(*
SPDX-License-Identifier: MIT
License: https://opensource.org/license/mit
*)

(*!
<summary>Owns two ordered single-cycle tests for topology regressions.</summary>
<description>
Owns persistent child storage and fixed parent associations. Use in one task without reentry.
Children is borrowed and must not be modified by application code. Constructor callbacks are not used.
Regression tests may deliberately corrupt the exposed array between failed operations to inject topology faults.
</description>
*)

{attribute 'no_assign'}
{attribute 'no_explicit_call' := 'do not call this function block directly'}
FUNCTION_BLOCK PairTestGroup EXTENDS TOF_Testing.TestGroup<2>
VAR_STAT
	//! <summary>Class name shared by all instances of this function block.</summary>
	{attribute 'hide'}
	_ClassName : STRING := __POUNAME();
END_VAR
VAR
	{attribute 'hide'}
	{attribute 'init_namespace'}
	_NamespaceName : STRING;
END_VAR
VAR_OUTPUT
	//! <summary>First owned regression leaf.</summary>
	First : TestingProbe(name := "First", parent := THIS^);
	//! <summary>Second owned regression leaf.</summary>
	Second : TestingProbe(name := "Second", parent := THIS^);
END_VAR
VAR
	_Children : ARRAY [0.._ChildCount - 1] OF TOF_Testing.ITestElement :=
	[
		First,
		Second
	];
END_VAR

//! <summary>Borrows the concrete class name for the lifetime of this instance; callers must not modify it.</summary>
{attribute 'monitoring' := 'call'}
PROPERTY ClassName : REFERENCE TO STRING
GET
ClassName REF= _ClassName;
END_GET
END_PROPERTY

//! <summary>Borrows the compiler-initialized namespace; callers must not modify the returned reference.</summary>
{attribute 'monitoring' := 'call'}
PROPERTY NamespaceName : REFERENCE TO STRING
GET
NamespaceName REF= _NamespaceName;
END_GET
END_PROPERTY

//! <summary>Reports the complete concrete instance size, excluding separately allocated storage.</summary>
{attribute 'monitoring' := 'call'}
PROPERTY SelfSize : ULINT
GET
SelfSize := XSIZEOF(THIS^);
END_GET
END_PROPERTY

//! <summary>Borrows the fixed array of this concrete group; do not modify it.</summary>
{attribute 'monitoring' := 'call'}
PROPERTY Children : REFERENCE TO ARRAY [0.._ChildCount - 1] OF TOF_Testing.ITestElement
GET
Children REF= _Children;
END_GET
END_PROPERTY

END_FUNCTION_BLOCK

(* stored: Version 1.1.0.1
   POU PairTestGroup: Id {a9015fc1-901f-4262-a805-9e04c9552dae}, SpecialFunc None
   Property ClassName: Id {e0dff1e8-c92d-4d74-b9a0-992c3919f486}
   Get Get: Id {ded61dfe-1470-4996-82a4-84727881dc42}
   Property NamespaceName: Id {8249691d-9f58-416a-adfc-84556791ffb0}
   Get Get: Id {de7120d0-a048-4428-a092-24eac5a85f37}
   Property SelfSize: Id {9c42e75d-9aa2-4202-80a3-7e5d37e006cd}
   Get Get: Id {d428cfff-8011-421e-a227-7739abac07fe}
   Property Children: Id {8b040fe0-48e4-4078-b98e-9ea7694ce02f}
   Get Get: Id {b0f2969f-6d03-47e7-a39a-779aab512d4b} *)
